(* IEC 61131-3 sources: trust-platform/libraries/plant/examples/sequences/src, 3 files *)

(* ---- FillSequence.st ---- *)
(* A customer sequence: fill a tank to a target level, hold it there for a mixing time, then drain
   it. Hold pauses with the valves closed and the timer standing still; Stop drains the tank before
   it ends. The manager overview needs no change for a new sequence. *)
USING Plant;

FUNCTION_BLOCK FillSequence EXTENDS Plant.FB_Sequence
VAR_INPUT
    Level : LREAL;
    TargetLevel : LREAL := 2.0;
    EmptyLevel : LREAL := 0.1;
    MixingTime : TIME := T#5m;
END_VAR
VAR_OUTPUT
    OpenInlet : BOOL;
    OpenOutlet : BOOL;
    RunMixer : BOOL;
END_VAR
    OpenInlet := FALSE;
    OpenOutlet := FALSE;
    RunMixer := FALSE;
    IF Execute() THEN
        CASE CurrentStep OF
            0:
                GoTo(Number := 10, Name := 'Fill');
            10:
                OpenInlet := TRUE;
                Wait(Text := 'Filling to the target level');
                IF Level >= TargetLevel THEN
                    GoTo(Number := 20, Name := 'Mix');
                ELSE
                    StepTimeout(Limit := T#30m, Text := 'The tank did not fill within 30 min');
                END_IF;
            20:
                RunMixer := TRUE;
                IF StepTime >= MixingTime THEN
                    GoTo(Number := 30, Name := 'Drain');
                END_IF;
            30:
                OpenOutlet := TRUE;
                IF Level <= EmptyLevel THEN
                    Complete();
                ELSE
                    StepTimeout(Limit := T#30m, Text := 'The tank did not drain within 30 min');
                END_IF;
        END_CASE;
    ELSIF State = E_SequenceState#Stopping THEN
        OpenOutlet := TRUE;
        Wait(Text := 'Draining before stopping');
        IF Level <= EmptyLevel THEN
            StopDone();
        END_IF;
    END_IF;
END_FUNCTION_BLOCK

(* ---- Configuration.st ---- *)
CONFIGURATION Tanks
RESOURCE Cpu ON PLC
    TASK Process (INTERVAL := T#100ms, PRIORITY := 1);
    PROGRAM Plant1 WITH Process : Main;
END_RESOURCE
END_CONFIGURATION

(* ---- Main.st ---- *)
(* Two tanks, each filled by its own FillSequence; one FB_SequenceManager shows both and can stop
   them together. Valves and mixers are Plant devices commanded in Auto by the sequences. *)
USING Plant;

PROGRAM Main
VAR
    Level1Signal : LREAL;
    Level2Signal : LREAL;
    Inlet1Out : BOOL;
    Outlet1Out : BOOL;
    Inlet2Out : BOOL;
    Outlet2Out : BOOL;
    Mixer1Out : BOOL;
    Mixer2Out : BOOL;

    Level1 : Plant.FB_LevelInput := (Unit := 'm', RangeHigh := 3.0);
    Level2 : Plant.FB_LevelInput := (Unit := 'm', RangeHigh := 3.0);
    Inlet1 : Plant.FB_OnOffValve := (HasOpenFeedback := FALSE, HasClosedFeedback := FALSE);
    Outlet1 : Plant.FB_OnOffValve := (HasOpenFeedback := FALSE, HasClosedFeedback := FALSE);
    Inlet2 : Plant.FB_OnOffValve := (HasOpenFeedback := FALSE, HasClosedFeedback := FALSE);
    Outlet2 : Plant.FB_OnOffValve := (HasOpenFeedback := FALSE, HasClosedFeedback := FALSE);
    Mixer1 : Plant.FB_Agitator := (HasFeedback := FALSE);
    Mixer2 : Plant.FB_Agitator := (HasFeedback := FALSE);
    Fill1 : FillSequence;
    Fill2 : FillSequence := (TargetLevel := 2.5);
    Overview : Plant.FB_SequenceManager;
END_VAR
    Level1(Raw := Level1Signal);
    Level2(Raw := Level2Signal);
    Fill1(Level := Level1.Value);
    Fill2(Level := Level2.Value);
    Overview(Sequence1 := Fill1, Sequence2 := Fill2);
    Inlet1(AutoOpen := Fill1.OpenInlet);
    Outlet1(AutoOpen := Fill1.OpenOutlet);
    Mixer1(AutoRun := Fill1.RunMixer);
    Inlet2(AutoOpen := Fill2.OpenInlet);
    Outlet2(AutoOpen := Fill2.OpenOutlet);
    Mixer2(AutoRun := Fill2.RunMixer);
    Inlet1Out := Inlet1.Solenoid;
    Outlet1Out := Outlet1.Solenoid;
    Mixer1Out := Mixer1.RunCommand;
    Inlet2Out := Inlet2.Solenoid;
    Outlet2Out := Outlet2.Solenoid;
    Mixer2Out := Mixer2.RunCommand;
END_PROGRAM
